Fanuc KAREL source: KD00058.KL

PROGRAM KD00058
%NOLOCKGROUP
VAR
  I: INTEGER
  J: INTEGER
  B: BOOLEAN
  R: REAL
  S: STRING[80]
BEGIN
  CONDITION[1]:
  WHEN DIN[1] = ON DO
    ABORT
  ENDCONDITION
END KD00058
